// TIA Portal V18 export
TYPE "UDT_EquipamentoScala"
   STRUCT
      Equipamento : Array[1..18] of "UDT_DadosEquipScala";
   END_STRUCT;
END_TYPE
